FUNCTION_BLOCK _TcVnMatrix3x3_LREAL_TestSuite EXTENDS TcUnit.FB_TestSuite
VAR
END_VAR

TestTryDeserializeFromNested();
TestTryDeserializeFromFlat();
TestTryDeserializeFromMixedFails();
TestTryDeserializeFromBadElementFails();
TestTryDeserializeFromFlat2x3();

METHOD PUBLIC TestTryDeserializeFromNested
VAR
    deserializer : JsonDeserializer;
    feedback : DeserializerFeedback;
    json : STRING(255) := '[[1,2,3],[4,5,6],[7,8,9]]';
    _type : _TcVnMatrix3x3_LREAL;
    result : BOOL;
END_VAR
TEST('TestTryDeserializeFromNested');

deserializer.Reset();
deserializer.TryLoad(json);
result := _type.TryDeserializeFrom(deserializer, feedback);

AssertTrue(Condition := result, Message := 'Deserialization reported failure.');
AssertEquals_LREAL(Expected := 2, Actual := _type.Value[0, 1], Delta := 0.0, Message := 'Nested value: [0, 1] wrong (row-major order expected).');
AssertEquals_LREAL(Expected := 4, Actual := _type.Value[1, 0], Delta := 0.0, Message := 'Nested value: [1, 0] wrong (row-major order expected).');
AssertEquals_LREAL(Expected := 9, Actual := _type.Value[2, 2], Delta := 0.0, Message := 'Nested value: [2, 2] wrong.');

TEST_FINISHED();
END_METHOD

METHOD PUBLIC TestTryDeserializeFromFlat
VAR
    deserializer : JsonDeserializer;
    feedback : DeserializerFeedback;
    json : STRING(255) := '[1,2,3,4,5,6,7,8,9]';
    _type : _TcVnMatrix3x3_LREAL;
    result : BOOL;
END_VAR
TEST('TestTryDeserializeFromFlat');

deserializer.Reset();
deserializer.TryLoad(json);
result := _type.TryDeserializeFrom(deserializer, feedback);

AssertTrue(Condition := result, Message := 'Deserialization reported failure.');
AssertEquals_LREAL(Expected := 2, Actual := _type.Value[0, 1], Delta := 0.0, Message := 'Flat value: [0, 1] wrong (row-major order expected).');
AssertEquals_LREAL(Expected := 4, Actual := _type.Value[1, 0], Delta := 0.0, Message := 'Flat value: [1, 0] wrong (row-major order expected).');
AssertEquals_LREAL(Expected := 9, Actual := _type.Value[2, 2], Delta := 0.0, Message := 'Flat value: [2, 2] wrong.');

TEST_FINISHED();
END_METHOD

METHOD PUBLIC TestTryDeserializeFromMixedFails
VAR
    deserializer : JsonDeserializer;
    feedback : DeserializerFeedback;
    json : STRING(255) := '[1,2,3,[4,5,6],7,8,9]';
    _type : _TcVnMatrix3x3_LREAL;
    result : BOOL;
END_VAR
TEST('TestTryDeserializeFromMixedFails');

deserializer.Reset();
deserializer.TryLoad(json);
result := _type.TryDeserializeFrom(deserializer, feedback);

AssertFalse(Condition := result, Message := 'A mix of flat and nested elements must fail.');

TEST_FINISHED();
END_METHOD

METHOD PUBLIC TestTryDeserializeFromBadElementFails
VAR
    deserializer : JsonDeserializer;
    feedback : DeserializerFeedback;
    json : STRING(255) := '[1,2,"x",4,5,6,7,8,9]';
    _type : _TcVnMatrix3x3_LREAL;
    result : BOOL;
END_VAR
TEST('TestTryDeserializeFromBadElementFails');

deserializer.Reset();
deserializer.TryLoad(json);
result := _type.TryDeserializeFrom(deserializer, feedback);

AssertFalse(Condition := result, Message := 'A non-numeric element must fail.');

TEST_FINISHED();
END_METHOD

METHOD PUBLIC TestTryDeserializeFromFlat2x3
VAR
    deserializer : JsonDeserializer;
    feedback : DeserializerFeedback;
    json : STRING(255) := '[1,2,3,4,5,6]';
    _type : _TcVnMatrix2x3_LREAL;
    result : BOOL;
END_VAR
TEST('TestTryDeserializeFromFlat2x3');

deserializer.Reset();
deserializer.TryLoad(json);
result := _type.TryDeserializeFrom(deserializer, feedback);

AssertTrue(Condition := result, Message := 'Deserialization reported failure.');
AssertEquals_LREAL(Expected := 3, Actual := _type.Value[0, 2], Delta := 0.0, Message := 'Flat 2x3 value: [0, 2] wrong.');
AssertEquals_LREAL(Expected := 4, Actual := _type.Value[1, 0], Delta := 0.0, Message := 'Flat 2x3 value: [1, 0] wrong (row-major order expected).');
AssertEquals_LREAL(Expected := 6, Actual := _type.Value[1, 2], Delta := 0.0, Message := 'Flat 2x3 value: [1, 2] wrong.');

TEST_FINISHED();
END_METHOD

END_FUNCTION_BLOCK

(* stored: Version 1.1.0.1, ProductVersion 3.1.4024.13
   POU _TcVnMatrix3x3_LREAL_TestSuite: Id {28e0044d-9112-403d-b424-4530a9577957}, SpecialFunc None
   Method TestTryDeserializeFromNested: Id {7bb3d6a9-c7b6-49f1-bb00-c2b1f3e985dd}
   Method TestTryDeserializeFromFlat: Id {63ba3579-1d67-484e-ad4e-69a7a2e3d114}
   Method TestTryDeserializeFromMixedFails: Id {eb565c5a-4fe7-4921-af56-4257942cf242}
   Method TestTryDeserializeFromBadElementFails: Id {d1016fd6-c774-40e8-843c-91ee0cdcd04f}
   Method TestTryDeserializeFromFlat2x3: Id {2c71a6fd-2958-44ae-9f1d-e2abff88f108} *)
